RoboDK station: animacion root.rdk

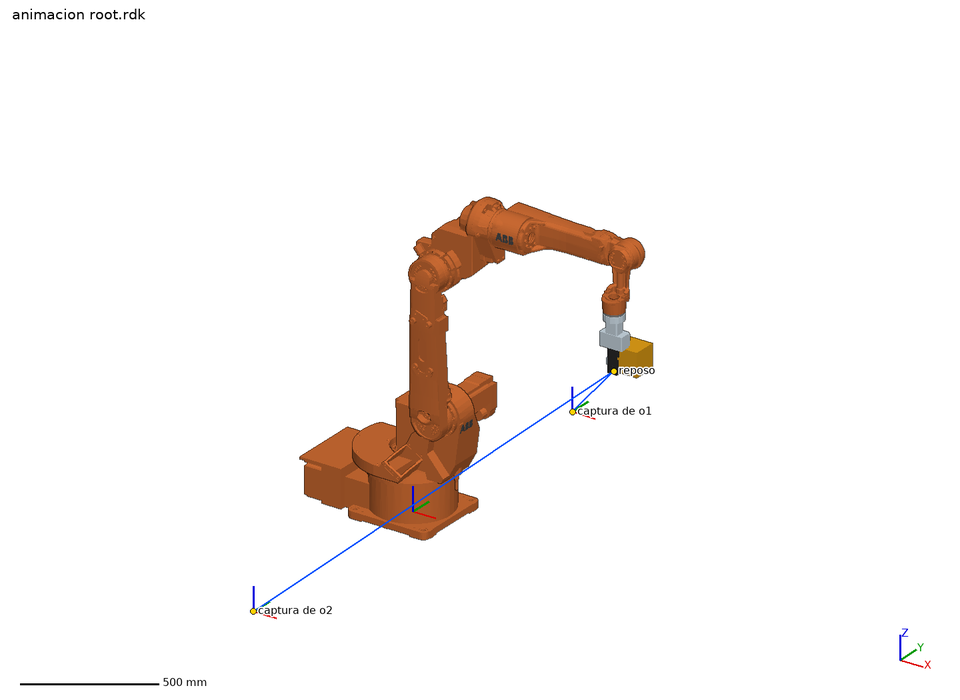
[picture v0: the station drawn from its stored meshes, robots at their saved joint values, targets as dots, program paths as lines]
Station animacion root (saved by RoboDK 5.6.5). Poses are relative to the parent item; angles as X-Y-Z fixed-axis rotations.
  - frame ABB IRB 1520ID Base at (0, 0, 0) mm
    - robot ABB IRB 1520ID: 6 axes, payload 5 kg, reach 1450 mm, repeatability 0.05 mm, weight 170 kg
        modified DH rows (alpha deg, a mm, theta deg, d mm): 0, 0, 0, 453; -90, 160, -90, 0; 0, 590, 0, 0; -90, 200, 0, 723; 90, 0, 0, 0; -90, 0, 180, 200
        joint limits [-170, -90, -100, -155, -135, -200] to [170, 150, 80, 155, 135, 200]; home [0, 0, 0, 0, 0, 0]; saved at [0, 0, 0, 0, 90, 0]
      - tool Generic 2-Finger Gripper, TCP at (0, 0, 233.37) mm, size 100 x 89.2 x 240.5 mm
        - object Cube 100mm at (0, 0, 0) mm, rotated rx 180 ry 0 rz -180 deg, size 100 x 100 x 100 mm, geometry from Cube-100mm.sld
  - frame Posicion 1 at (0, 1000, 0) mm
    - target reposo (Cartesian target) at (883, -1000, 809.63) mm, rotated rx 180 ry 0 rz -180 deg; joints [0, 0, 0, 0, 90, 0] of ABB IRB 1520ID
    - target captura de o1 (Cartesian target) at (0, 0, 0) mm, rotated rx 180 ry 0 rz -180 deg; joints [90, 31.047, 28.843, 0, 30.11, 90] of ABB IRB 1520ID
    - target captura de o2 (Cartesian target) at (0, -2000.86, 0) mm, rotated rx 180 ry 0 rz -180 deg; joints [-90, 31.108, 28.747, 0, 30.145, -90] of ABB IRB 1520ID
    - target Target 4 (Cartesian target) at (0, -2000.86, 0) mm, rotated rx 180 ry 0 rz -180 deg; joints [-90, 31.108, 28.747, 0, 30.145, -90] of ABB IRB 1520ID
    - target Target 5 (Cartesian target) at (0, -2000.86, 0) mm, rotated rx 180 ry 0 rz -180 deg; joints [-90, 31.108, 28.747, 0, 30.145, -90] of ABB IRB 1520ID
    - target Target 6 (Cartesian target) at (0, -2000.86, 0) mm, rotated rx 180 ry 0 rz -180 deg; joints [-90, 31.108, 28.747, 0, 30.145, -90] of ABB IRB 1520ID
    - target Target 7 (Cartesian target) at (0, -2000.86, 0) mm, rotated rx 180 ry 0 rz -180 deg; joints [-90, 31.108, 28.747, 0, 30.145, -90] of ABB IRB 1520ID
    - target Target 8 (Cartesian target) at (0, -2000.86, 0) mm, rotated rx 180 ry 0 rz -180 deg; joints [-90, 31.108, 28.747, 0, 30.145, -90] of ABB IRB 1520ID
    - target Target 9 (Cartesian target) at (883, -1000, 809.63) mm, rotated rx 180 ry 0 rz -180 deg; joints [0, 0, 0, 0, 90, 0] of ABB IRB 1520ID
    - target Target 10 (Cartesian target) at (883, -1000, 809.63) mm, rotated rx 180 ry 0 rz -180 deg; joints [0, 0, 0, 0, 90, 0] of ABB IRB 1520ID
    - target Target 11 (Cartesian target) at (883, -1000, 809.63) mm, rotated rx 180 ry 0 rz -180 deg; joints [0, 0, 0, 0, 90, 0] of ABB IRB 1520ID
    - target Target 12 (Cartesian target) at (883, -1000, 809.63) mm, rotated rx 180 ry 0 rz -180 deg; joints [0, 0, 0, 0, 90, 0] of ABB IRB 1520ID
  - frame Posicion 2 at (0, -1000.86, 0) mm
  - program Prog1 (15 instructions, listed below)
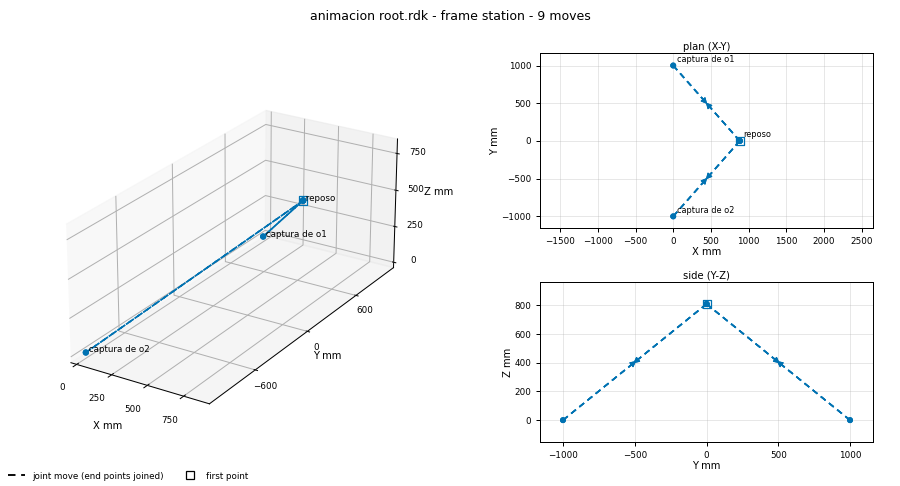
[picture p0: tool path of animacion root.rdk in frame station, 9 of 9 moves have a stored position in this frame; points joined in program order, loops and branches not executed]

--- program Prog1 (robot ABB IRB 1520ID) ---
  Est. Ref.: Posicion 1
  Est. herr: Generic 2-Finger Gripper
  MoveJ (reposo)
  MoveJ (captura de o1)
  Adjuntar a Generic 2-Finger Gripper
  MoveJ (reposo)
  MoveJ (captura de o2)
  Separar de Generic 2-Finger Gripper
  MoveJ (reposo)
  MoveJ (captura de o2)
  Adjuntar a Generic 2-Finger Gripper
  MoveJ (reposo)
  MoveJ (captura de o1)
  Separar de Generic 2-Finger Gripper
  MoveJ (reposo)
